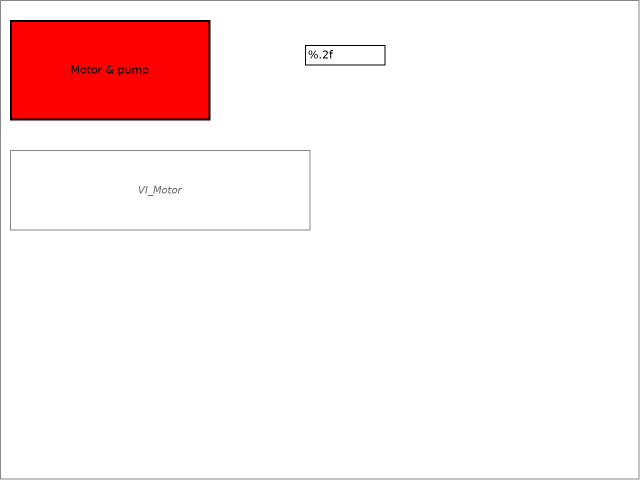
VISUALIZATION VI_Demo  // 640x480
VAR_IN_OUT
	fbMotor : FB_Motor;
END_VAR
    Rectangle (10,20 200x100), "Motor & pump"
    Group (300,40 100x40)
        Textfield (5,5 80x20), "%.2f", text variable: fbMotor.rSpeed
            OnMouseClick: write fbMotor.rSetSpeed via Default, min 0
    Frame (10,150 300x80)
        shows VI_Motor(fbMotor := MAIN.fbMotor1)
END_VISUALIZATION

(* stored: Version 1.1.0.1, ProductVersion 3.1.4024.12
   Visu VI_Demo: Id {11111111-2222-3333-4444-555555555555} *)
